// TIA Portal V21 export
DATA_BLOCK "IDB_FbdBoxes"   // DB22
// stored: InstanceOfName FB_FbdBoxes, InstanceOfType FB
"FB_FbdBoxes"
   // VAR_INPUT
   //    Start : Bool;
   //    InValue : Int;
   //    Limit : Int;
   // END_VAR
   // VAR_OUTPUT
   //    Delayed : Bool;
   //    Copy : Int;
   //    Sum : Int;
   //    IsEqual : Bool;
   //    SectionsOk : Bool;
   //    Skipped : Bool;
   //    AfterJump : Bool;
   // END_VAR
   // VAR
   //    Delay { S7_SetPoint := 'True'} : TON_TIME;
   //    DelayElapsed : Time;
   //    Timers { S7_SetPoint := 'True'} : "FB_SclTimers";
   //    TimerRunOn : Bool;
   //    TimerPulse : Bool;
   //    TimerCount : Int;
   //    TimerDelayed : Bool;
   //    TimerReached : Bool;
   // END_VAR
BEGIN
END_DATA_BLOCK
